FUNCTION_BLOCK ALARM_DEBOUNCE (* Migrated from IEC 61131-3 ST *)
  (* Standard: 61499-2 *)
  (* Version 1.0, 2026-11-06, st2fb *)
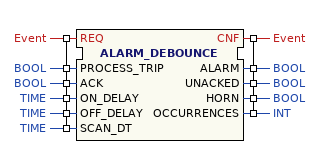
  EVENT_INPUT
    REQ WITH PROCESS_TRIP, ACK, ON_DELAY, OFF_DELAY, SCAN_DT;
  END_EVENT
  EVENT_OUTPUT
    CNF WITH ALARM, UNACKED, HORN, OCCURRENCES;
  END_EVENT
  VAR_INPUT
    PROCESS_TRIP : BOOL;
    ACK : BOOL;
    ON_DELAY : TIME;
    OFF_DELAY : TIME;
    SCAN_DT : TIME;
  END_VAR
  VAR_OUTPUT
    ALARM : BOOL;
    UNACKED : BOOL;
    HORN : BOOL;
    OCCURRENCES : INT;
  END_VAR
  VAR
    ST2FB_NOW : TIME := T#0s;
    ON_TIMER_IN : BOOL;
    ON_TIMER_PT : TIME := T#0s;
    ON_TIMER_Q : BOOL;
    ON_TIMER_ET : TIME := T#0s;
    ON_TIMER_STATE : INT := 0;
    ON_TIMER_PREV_IN : BOOL;
    ON_TIMER_START_TIME : TIME := T#0s;
    OFF_TIMER_IN : BOOL;
    OFF_TIMER_PT : TIME := T#0s;
    OFF_TIMER_Q : BOOL;
    OFF_TIMER_ET : TIME := T#0s;
    OFF_TIMER_STATE : INT := 0;
    OFF_TIMER_PREV_IN : BOOL;
    OFF_TIMER_START_TIME : TIME := T#0s;
    RAISED_CLK : BOOL;
    RAISED_Q : BOOL;
    RAISED_M : BOOL;
    ACK_EDGE_CLK : BOOL;
    ACK_EDGE_Q : BOOL;
    ACK_EDGE_M : BOOL;
  END_VAR
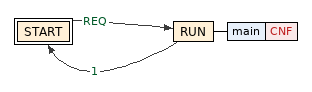
  EC_STATES
    START;
    RUN : main -> CNF;
  END_STATES
  EC_TRANSITIONS
    START TO RUN := REQ;
    RUN TO START := 1;
  END_TRANSITIONS
  ALGORITHM main IN ST:
ST2FB_NOW := ST2FB_NOW + SCAN_DT;

ON_TIMER_IN := PROCESS_TRIP;
ON_TIMER_PT := ON_DELAY;
IF (ON_TIMER_STATE = 0) AND NOT ON_TIMER_PREV_IN AND ON_TIMER_IN THEN
  ON_TIMER_STATE := 1;
  ON_TIMER_Q := FALSE;
  ON_TIMER_START_TIME := ST2FB_NOW;
ELSE
  IF NOT ON_TIMER_IN THEN
    ON_TIMER_ET := T#0s;
    ON_TIMER_Q := FALSE;
    ON_TIMER_STATE := 0;
  ELSIF ON_TIMER_STATE = 1 THEN
    IF ON_TIMER_START_TIME + ON_TIMER_PT <= ST2FB_NOW THEN
      ON_TIMER_STATE := 2;
      ON_TIMER_Q := TRUE;
      ON_TIMER_ET := ON_TIMER_PT;
    ELSE
      ON_TIMER_ET := ST2FB_NOW - ON_TIMER_START_TIME;
    END_IF;
  END_IF;
END_IF;
ON_TIMER_PREV_IN := ON_TIMER_IN;

OFF_TIMER_IN := ON_TIMER_Q;
OFF_TIMER_PT := OFF_DELAY;
IF (OFF_TIMER_STATE = 0) AND OFF_TIMER_PREV_IN AND NOT OFF_TIMER_IN THEN
  OFF_TIMER_STATE := 1;
  OFF_TIMER_START_TIME := ST2FB_NOW;
ELSE
  IF OFF_TIMER_IN THEN
    OFF_TIMER_ET := T#0s;
    OFF_TIMER_STATE := 0;
  ELSIF OFF_TIMER_STATE = 1 THEN
    IF OFF_TIMER_START_TIME + OFF_TIMER_PT <= ST2FB_NOW THEN
      OFF_TIMER_STATE := 2;
      OFF_TIMER_ET := OFF_TIMER_PT;
    ELSE
      OFF_TIMER_ET := ST2FB_NOW - OFF_TIMER_START_TIME;
    END_IF;
  END_IF;
END_IF;
OFF_TIMER_Q := OFF_TIMER_IN OR (OFF_TIMER_STATE = 1);
OFF_TIMER_PREV_IN := OFF_TIMER_IN;

ALARM := OFF_TIMER_Q;

RAISED_CLK := ALARM;
RAISED_Q := RAISED_CLK AND NOT RAISED_M;
RAISED_M := RAISED_CLK;

ACK_EDGE_CLK := ACK;
ACK_EDGE_Q := ACK_EDGE_CLK AND NOT ACK_EDGE_M;
ACK_EDGE_M := ACK_EDGE_CLK;

IF RAISED_Q THEN
  UNACKED := TRUE;
  OCCURRENCES := OCCURRENCES + 1;
ELSIF ACK_EDGE_Q THEN
  UNACKED := FALSE;
END_IF;
HORN := ALARM AND UNACKED;
  END_ALGORITHM
END_FUNCTION_BLOCK
